Fanuc KAREL source: KT00784.KL

PROGRAM KT00784
%NOLOCKGROUP
VAR
  I1: INTEGER
  I2: INTEGER
  OUT: INTEGER
BEGIN
  I1 = 2
  I2 = 3
  I1 = 2
  I2 = 3
  OUT = COS(I1)
END KT00784
